(* IEC 61131-3 sources: test/Class/SafetyBaseFSoE (part 5) *)

      pSafetyManagerThis^.NewInst(#MyPara, #MyResult);

      QuitComError := MyResult.aData[0]$DINT;

      // refresh the server on the outer object
      RefreshAsySrv();
    end_if;

    // if we are reinitializing and we have a valid safety number
    if (SafetyState = _ReinitConfig) & SafetyNumber then

      // check every 3 seconds if the cpu is configured
      if b_CheckConfigured & ((ops.tAbsolute - ud_LastCheckConfig) > 3000) then

        // get state via SDO communication
        sd_retval := SDOStdRequ ( us_Command      := SBF_SDO_COMMAND_GET_STATE
                                , p_us_RespData   := ( #GetStateResp )$^USINT
                                , us_RespLength   := sizeof(GetStateResponseType)
                                );

        // the cpu is configured, load the new configuration
        if ( sd_retval = 0 ) &
           (GetStateResp.ConfigState <> SBF_CFG_STATE_UNKNOWN) &
           (GetStateResp.ConfigState <> SBF_CFG_STATE_INVALID) &
           (GetStateResp.ConfigState <> SBF_CFG_STATE_NOT_CONFIGURED) then

          b_CheckConfigured := FALSE;

          b_GetNewConfiguration := TRUE;
        end_if;

        // remember the last time we checked for configurated cpu
        ud_LastCheckConfig := ops.tAbsolute;
      end_if;

      // if there is a new configuration => get it
      if b_GetNewConfiguration then
        // get configuration from safe CPU and build routing tables
        sd_retval := GetRoutingData();
        if sd_retval = 0 then
          b_GetNewConfiguration := FALSE;

          SendAllUnsafeValues();
        else
          LogError("@024B (SafetyBaseFSoE::Background) FAILED TO REINIT THE SAFECPU: .");
        end_if;
      end_if;
    elsif ConnectionInfos.ConnectionNo then
      // if there are still connections => check if they are initialized
      CheckFSoEConnections();
    end_if;

    // here we save the log file from the module to the harddrive (started by user)
    if DiagVars.SavingLogInProgress then

      case DiagVars.SavingLogSSW of

  // ********************************************************************************************************************************************
        GetLogHeader:     // get log header from module (contains size of log memory and write counter)

          // get log header via SDO communication
          sd_retval := SDORequ ( us_Command      := SBF_SDO_COMMAND_GET_LOG_HDR
                               , p_us_RequData   := #DiagVars.ucChoiceSaveLog
                               , us_RequLength   := 1
                               , p_us_RespData   := ( #DiagVars.LogHeader)$^USINT
                               , us_RespLength   := sizeof(DiagStructType.LogHeader)
                               );

          if ( sd_retval = 0 ) then
            DiagVars.LogMemToGet := DiagVars.LogHeader.LogMemSize;
            DiagVars.pLogFileMem$pVoid := ToStdLib.Malloc(size:=DiagVars.LogHeader.LogMemSize);
            //_memset(dest:=DiagVars.pLogFileMem$pVoid, usByte:=0, cntr:=DiagVars.LogHeader.LogMemSize);
            if DiagVars.ucChoiceSaveLog = 0 then
              DiagVars.ReadBaseAdr := SBF_SDO_ADDRESS_LOG_UC1;
            else
              DiagVars.ReadBaseAdr := SBF_SDO_ADDRESS_LOG_UC2;
            end_if;
            DiagVars.SavingLogSSW := GetLogFileBlocks;

          end_if;

  // ********************************************************************************************************************************************
        GetLogFileBlocks: // get the log memory from the application memory of the module (every cycle only a little bit to prevent runtime error in module)

          // we wait here until UpdateCy finishes our work

  // ********************************************************************************************************************************************
        GetLogHeader2:    // get log header from module again. if write counter changed,
                          // we repeat GetLogFileBlocks. otherwise we continue to save the file

          LastWriteCounter := DiagVars.LogHeader.WriteCounter;

          // get LogHeader
          sd_retval := SDORequ ( us_Command      := SBF_SDO_COMMAND_GET_LOG_HDR
                               , p_us_RequData   := #DiagVars.ucChoiceSaveLog
                               , us_RequLength   := 1
                               , p_us_RespData   := ( #DiagVars.LogHeader)$^USINT
                               , us_RespLength   := sizeof(DiagStructType.LogHeader)
                               );

          if ( sd_retval = 0 ) then

            // if write counter is different, repeat last step
            if DiagVars.LogHeader.WriteCounter <> LastWriteCounter then
              DiagVars.SavingLogSSW := GetLogFileBlocks;

              DiagVars.LogMemToGet := DiagVars.LogHeader.LogMemSize;

              // realloc memory (maybe it's a different size)
              ToStdLib.Free(mptr:=DiagVars.pLogFileMem$pVoid);
              DiagVars.pLogFileMem$pVoid := ToStdLib.Malloc(size:=DiagVars.LogHeader.LogMemSize);
            else
              // write counter is equal. continue to last step
              DiagVars.SavingLogSSW := SaveLogFile;
            end_if;
          end_if;

  // ********************************************************************************************************************************************
        SaveLogFile:      // save the memory to the specified file (DPNE)

          // open file (create/overwrite always)
          FileHandle := FileSys.FileOpen(filename:=#DiagVars.DPNE[0], attributes:=ATT_CREATE_ALWAYS);

          DiagVars.SavingLogSuccessful := 1;

          if FileHandle >= 0 then

            // save content to it
            if FileSys.FileWrite(handle:=FileHandle, buffer:=DiagVars.pLogFileMem, length:=DiagVars.LogHeader.LogMemSize) <> DiagVars.LogHeader.LogMemSize$DINT then
              // failed to write to file
              LogError("@024C (SafetyBaseFSoE::Background) Failed to write to binary LogFile.");
              DiagVars.SavingLogSuccessful := -1;
            end_if;

            // close file
            FileSys.FileClose(handle:=FileHandle);
          else
            // failed to open file
            LogError("@024D (SafetyBaseFSoE::Background) Failed to open binary LogFile.");
            DiagVars.SavingLogSuccessful := -1;
          end_if;

          ToStdLib.Free(mptr:=DiagVars.pLogFileMem$pVoid);
          DiagVars.pLogFileMem := NIL;

          DiagVars.SavingLogSSW := GetLogHeader;
          DiagVars.SavingLogInProgress := FALSE;

      end_case;
    end_if;
  end_if;

  state := READY;

END_FUNCTION

FUNCTION VIRTUAL GLOBAL SafetyBaseFSoE::RtWork
  VAR_INPUT
    EAX 	: UDINT;
  END_VAR
  VAR_OUTPUT
    state (EAX) 	: UDINT;
  END_VAR
  VAR
    calloption    : UDINT;
    PDOLength     : UINT;
    pBuffer       : ^USINT;
    pDOInfo       : ^t_DOInfo;
    i             : USINT;
  END_VAR

  // Save state
  // This must be the 1. line in this function or EAX may be overwritten by the generated AWL code
  calloption := EAX;

  if calloption = CALL_OPTION_RT_PRESCAN then    // Called from UpdateRt

//============================ Profiler start======================================================
#ifdef  DM_Profiler
    StartTimeMeasurement(usMode := DMTIME_RT);
#endif
//============================ Profiler end========================================================

    // do pdo communication only, if module has been found and initialized correctly and if there are some LEDs on (else a FW-Update is running)
    if Online &
       (( SafetyState = _SafetyClassOK ) | ( SafetyState = _WaitForSynchronicity ) | ( SafetyState = _ReinitConfig ) | ( SafetyState = _ModFromCfgNotFound ) | ( SafetyState = _UnknownCfgError ) | ( SafetyState = _UnsafeVarNotFound )) then

      // get I/O state, runstate, error
      UpDateNotStd(calloption:=calloption);

      // wait until the safetymanager has initialized everything
      if b_ManagerInitialisationFinished = FALSE then
        return;
      end_if;

      // if any LED is active, then firmware update is not active and we can do our work
      if (VoltageOK | RunState | ServiceMode | ErrorState) then
        // if we are in run state
        if RunState then
          if PDOSingleRunActive & WriteDOsUsed then
            PDOSingleRunActive -= 1;
            if PDOSingleRunActive = 0 then
              for i := 0 to WriteDOsUsed-1 do
                SetDORunState(Handle:=aWritePDOs[i].Handle, NewState:=_BUS_IF_RUN_STATE_NO_RUN);
              end_for;
            end_if;
          end_if;

          //read PDO from hardware, only if PDO is needed by other moduls
          if ( PDOOutputIsUsed ) & ReadDOsUsed then

            PDOLength := pPDOLengthInfoData^.PDOReadLength;

            // only if length is bigger than minimum and smaller than maximum
            if ( PDOLength >= SBF_SPDO_MIN_LENGTH ) & ( PDOLength <= MyPDOReadSize) then

              pBuffer := #PDOOutputBuffer[0];
              pDOInfo := #aReadPDOs[0];
              for i := 0 to (ReadDOsUsed-1) do
                _memcpy(ptr1:=pBuffer, ptr2:=pDOInfo^.pData, cntr:=pDOInfo^.Length);
                pBuffer += pDOInfo^.Length;
                pDOInfo += sizeof(t_DOInfo);
              end_for;

#ifdef SAFETY_PROTOCOL_ANALYZER_ACTIVATED
  RecordFrame(pFrame:=(#PDOOutputBuffer[0])$^DINT, FrameState:=0, IsFSoEPDO:=TRUE);
#endif
            else
              InvalidPDOSizeCnt += 1;
            end_if;
          end_if;
        end_if;
      end_if;
    end_if;

//============================ Profiler start======================================================
#ifdef  DM_Profiler
    StopTimeMeasurement(usMode := DMTIME_RT);
#endif
//============================ Profiler end========================================================

  elsif calloption = CALL_OPTION_RT_POSTSCAN then // Called from UpdateRtPostScan

//============================ Profiler start======================================================
#ifdef  DM_Profiler
    StartTimeMeasurement(usMode := DMTIME_RTPOSTSCAN);
#endif
//============================ Profiler end========================================================

    // do pdo communication only, if module has been found and initialized correctly and if there are some LEDs on (else a FW-Update is running)
    if Online &
       (( SafetyState = _SafetyClassOK ) | ( SafetyState = _WaitForSynchronicity ) | ( SafetyState = _ModFromCfgNotFound ) | ( SafetyState = _UnknownCfgError ) | ( SafetyState = _UnsafeVarNotFound )) then

      // if any LED is active, then firmware update is not active and we can do our work
      if (VoltageOK | RunState | ServiceMode | ErrorState) then

        // write unsafe I/Os
        UpDateNotStd(calloption:=calloption);

        if RunState & ((us_SetBusReadyState = SetBusReadyFinished) | b_ManualQuit) then
          //write PDO to hardware
          if ( ui_cnt_PDOInputBuffer > 0 ) then
            WritePDO2Module();
          end_if;
        end_if;
      end_if;
    end_if;

//============================ Profiler start======================================================
#ifdef  DM_Profiler
    StopTimeMeasurement(usMode := DMTIME_RTPOSTSCAN);
#endif
//============================ Profiler end========================================================
  end_if;

  state := READY;

END_FUNCTION

FUNCTION VIRTUAL GLOBAL SafetyBaseFSoE::ConnectEvent
  VAR
    MyPara 	              : CmdStruct;
    MyResult	            : results;
  END_VAR

  //start DOs
  StartDO();

  if SafetyState = _ModuleNotFound then
    if ModuleSyncNo = 0 then
      SetSafetyState(NewState:=_SafetyClassOK);
    else
      SetSafetyState(NewState:=_WaitForSynchronicity);
    end_if;
  end_if;

  // if we we're already connected => tell the sdias manager we're back (safetythis has to be valid if b_Reconnect is set, therefore we don't have to check it here)
  if b_Reconnect then
    MyPara.uiCmd := CMD_SM_MODULE_RECONNECT;
    MyPara.aPara[0] := THIS$DINT;
    pSafetyManagerThis^.NewInst(#MyPara, #MyResult);
  end_if;

  // whenever the postinit has passed and we got a connect (module has been plugged in after booting the application) => get it's config
  if b_PostInitPassed = TRUE then
    // start reading the config in background (if we're in init the post-init read-out will be faster)

    // next time we check for the configured state of the cpu
    b_CheckConfigured := TRUE;

    // check again in background
    SetSafetyState(NewState:=_ReinitConfig);
  end_if;

// online is set if module init succeeds
//  Online := 1;

END_FUNCTION

FUNCTION VIRTUAL GLOBAL SafetyBaseFSoE::DisconnectEvent
  VAR
    MyPara 	              : CmdStruct;
    MyResult	            : results;
  END_VAR

  //stop DOs
  StopDO();

  // reset time sync state and tell the manager
  if pSafetyManagerThis then
    MyPara.uiCmd := CMD_SM_MODULE_DISCONNECT;
    MyPara.aPara[0] := THIS$DINT;
    pSafetyManagerThis^.NewInst(#MyPara, #MyResult);

    b_Reconnect := TRUE;
  end_if;

  // clear request, otherwise problems could occur on next connect
  LastRequest := _NoOpenRequest;
  ud_AsyComRetryCounter := 0; // reset retry counter

  SafetyNumber := 0;
  FirmwareVersion := 0;

  // increment the config checksum to ensure the readout on reconnect (config readout also contains check of connected modules)
  DesignerPrjConfigCRC += 1;

  SetSafetyState(NewState:=_ModuleNotFound);

  // remove the cpu from all classes, which use it
  ResetConfig();

  if UnsafeScheduler <> UnsafeSchedulerSetBusReady then
    us_SetBusReadyState := WaitPDOsSyncron;
    UnsafeScheduler := UnsafeSchedulerSetBusReady;
  end_if;

  MaxVarsPerReadPackage := 0;
  ReadFramesNeeded := 0;
  MaxVarsPerWritePackage := 0;
  WriteFramesNeeded := 0;

  Online := 0;

END_FUNCTION

FUNCTION VIRTUAL GLOBAL SafetyBaseFSoE::InterruptEvent

END_FUNCTION

FUNCTION SafetyBaseFSoE::SetDORunState
  VAR_INPUT
    Handle 	: UDINT;
    NewState 	: t_BusIFRunState;
  END_VAR
  VAR
    dataSETRUNSTATE : t_SetRunStateCfg;
    tempCmd : CmdStruct;
    _result : results;
  END_VAR

  // set runstate of read
  dataSETRUNSTATE.Handle      := Handle;
  dataSETRUNSTATE.NewRunState := NewState;

  tempCmd.uiCmd         := _BUS_IF_SET_RUN_STATE;
  tempCmd.aPara[0]      := (#dataSETRUNSTATE)$DINT;

  ToBusInterface.NewInst(pPara:=#tempCmd, pResult:=#_result);

  if _result.aData[0]$t_BusIFRetvalErrorcode <> _BUS_IF_RETVAL_OK then
    if NewState = _BUS_IF_RUN_STATE_NO_RUN then
      DOStopFailCounter += 1;
    else
      DOStartFailCounter += 1;
    end_if;
  end_if;

END_FUNCTION

FUNCTION VIRTUAL GLOBAL SafetyBaseFSoE::CyWork
  VAR_INPUT
    EAX 	: UDINT;
  END_VAR
  VAR_OUTPUT
    state (EAX) 	: UDINT;
  END_VAR
  VAR
    p_SDO_act             : ^SDOHeader;
    us_SDO_length         : USINT;
    i                     : UINT;
    p_ReceiveObj          : pVirtualBase;
    p_SDOviaPath          : ^SDOviaPath;
    sd_retval             : DINT;
    IsStandardResp        : BOOL;
    SDORequestBuffer      : SDORequReadConfig;
    DataLen               : USINT;
    us_UnsafeSchedulerRun : USINT;
    p_PDOInBufferAct      : ^PDOInputBuffer;
    EverythingSynchron    : BOOL;
    MyPara 	              : CmdStruct;
    MyResult	            : results;
    UnsafeWrPackageNo     : USINT;
    aUnsafeWrPackages     : UnsafeWritePackages;
    UnsafeRdPackageNo     : USINT;
    aUnsafeRdPackages     : UnsafeReadPackages;
    TmpVal                : DINT;
    AddUnsafePackage      : BOOL;
    GotNewUnsafeValue     : BOOL;
    pHelpUnsafe           : ^UnsafeIORoutingElement;
    BDINTWriteVars        : USINT;
    pAddDynSlaveResp      : ^t_AddDynSlaveResponse;
  END_VAR

//============================ Profiler start======================================================
#ifdef  DM_Profiler
  StartTimeMeasurement(usMode := DMTIME_CY);
#endif
//============================ Profiler end========================================================

#ifdef HWK_SHOW_PRAGMA_MESSAGES
  if b_LogFirstDone = 1 then
    for i := 0 to (ui_cnt_PDOInputBuffer-1) do
      LogValue("@027F (SafetyBaseFSoE::WritePDO2Module) Copy 0x{0} Bytes to offset 0x{1} of Write PDO Nr. 0x{2}", Value:=aLogValues[i].ByteLen, Value2:=aLogValues[i].Offset, Value3:=aLogValues[i].DOIndex);
    end_for;

    b_LogFirstDone := 2;
  end_if;
#endif

  // do sdo communication only, if module has been found and initialized correctly and if there are some LEDs on (else a FW-Update is running)
  if Online & (VoltageOK | RunState | ServiceMode | ErrorState) &
     (( SafetyState <> _ModuleNotFound ) & ( SafetyState <> _MemAllocFailed ) & ( SafetyState <> _LostPowerSupply ) & ( SafetyState <> _ReadFWVerFailed ) & ( SafetyState <> _WrongSafetyHW ) & ( SafetyState <> _ReinitConfig )) then

    // wait until the safetymanager has initialized connection
    if (b_ManagerReadyForSDO = FALSE) then
      return;
    end_if;

    //Update of service messages doesn't take place in realtime

    //read SDO from module and send it to the target module
    //check, if SDO is available and valid
    if ( p_Handle_SDO_Read^.us_Status = SAFETY_SDO_DATA_VALID ) then

      //calculate length of SDO
      us_SDO_length := sizeof(SDOHeader.StdHeader.CRC) + p_Handle_SDO_Read^.SDOStructure.SDOHeader.StdHeader.Len;

      //copy SDO without first byte (=status byte)
      ToStdLib.MemCpy(dest := p_SDOOutputBuffer, source := #p_Handle_SDO_Read^.SDOStructure, size := us_SDO_length );

#ifdef SAFETY_PROTOCOL_ANALYZER_ACTIVATED
  RecordFrame(p_SDOOutputBuffer$^DINT, 0);
#endif

      //mark data as received
      p_Handle_SDO_Read^.us_Status := SAFETY_SDO_NO_DATA;

      //find target object for routing
      p_ReceiveObj := NIL;

      IsStandardResp := FALSE;
      //check, if receiver is addressed by safety number or hardware path
      if ((p_SDOOutputBuffer^.SDOHeader.StdHeader.Typ$USINT AND SBF_SSDO_MASK_TYPE)$t_SafetyFrameType = SSDO_MOD) then

        //search this-pointer of receiver with safety number
        p_ReceiveObj := ( GetRoutingPointerByNumber(ud_SafeNumber := p_SDOOutputBuffer^.SDOHeader.DstAdr))$pVirtualBase;

      elsif ((p_SDOOutputBuffer^.SDOHeader.StdHeader.Typ$USINT AND SBF_SSDO_MASK_TYPE)$t_SafetyFrameType = SSDO_MOD_TP) then

        //search this-pointer of receiver with hardware path
        p_SDOviaPath := p_SDOOutputBuffer$^SDOviaPath;
        p_ReceiveObj := ( GetRoutingPointerByPath(p_ActObjectPath := #p_SDOviaPath^.TopologyPath[0], p_SDOviaPath^.StdHeader.Len - 8))$pVirtualBase;
      elsif ((p_SDOOutputBuffer^.SDOHeader.StdHeader.Typ$USINT AND SBF_SSDO_MASK_TYPE)$t_SafetyFrameType = SDO_STD) then
        IsStandardResp := TRUE;
        StandardResponse := (p_SDOOutputBuffer$^StandardFrameType)^;
        if StandardResponse.SDOHeader.SeqNr = (StandardSeqNr OR 16#80) then

          // if the microcontroller got powered again and we have an SDO response => also get the configuration (don't wait the whole time)
          //if b_WaitForFirmwareBoot = TRUE then // no if to be faster (if it's false, it does not matter if we set it again to false)
          b_WaitForFirmwareBoot := FALSE;
          //end_if;

          case LastRequest of
            _NoOpenRequest: // error, no open request, but we got a response
              LogError("@0252 (SafetyBaseFSoE::CyWork) Standard frame response received, without open request.");

            _SetBusReady:
              IF StandardResponse.SDOHeader.Cmd = SBF_SDO_COMMAND_SET_BUS_READY THEN
                if us_SetBusReadyState <> SendSetBusReady then
                  LogError("@0253 (SafetyBaseFSoE::CyWork) Got Response of SetBusReady, but SSW is not in the right step.");
                  return;
                end_if;
                us_SetBusReadyState := SetBusReadyFinished;
                b_ManualQuit := FALSE;
                UnsafeScheduler := UnsafeSchedulerGetDiagVars; // Go on with the action-steps, done here so we don't lose a whole cycle
                LastRequest := _NoOpenRequest;
                ud_AsyComRetryCounter := 0; // reset retry counter
                if SafetyState = _WaitForSynchronicity then
                  SetSafetyState(NewState:=_SafetyClassOK);
                end_if;
              else
                LogError("@0256 (SafetyBaseFSoE::CyWork) Invalid command: bus ready expected.");
              END_IF;

            _ReadData:
              // if we did read command, then save the value to corresponding server
              if StandardResponse.SDOHeader.Cmd = SBF_SDO_COMMAND_READ then
                // if returncode is 0 read succeeded
                if StandardResponse.aData[0] = 0 then
                  // check if length is correct
                  if StandardResponse.aData[1] = StandardRequest.aData[4] then
                    // delete request
                    LastRequest := _NoOpenRequest;
                    ud_AsyComRetryCounter := 0; // reset retry counter

                    if (DiagVars.SavingLogSSW = GetLogFileBlocks) then
                      // save the last block in the memory for the file
                      _memcpy(ptr1:=DiagVars.pLogFileMem$pVoid + (DiagVars.LogHeader.LogMemSize - DiagVars.LogMemToGet),
                              ptr2:=#StandardResponse.aData[2],
                              cntr:=DiagVars.BytesToGet);

                      DiagVars.LogMemToGet -= DiagVars.BytesToGet;

                      if DiagVars.LogMemToGet = 0 then
                        DiagVars.SavingLogSSW := GetLogHeader2;
                      end_if;
                    else
                      LogError("@0255 (SafetyBaseFSoE::CyWork) SDO Receive: Invalid Read response (no diagnostic read active).");
                    end_if;
                  end_if;
                end_if;
              else
                LogError("@0256 (SafetyBaseFSoE::CyWork) SDO Receive: Invalid command, read expected.");
              end_if;

            _ReadValues:
              // if we did read command, then save the value to corresponding server
              if StandardResponse.SDOHeader.Cmd = SBF_SDO_COMMAND_READ_VALUES then
                // if returncode is 0 read succeeded
                if StandardResponse.aData[0] = 0 then
                  // check if length is correct
                  if StandardResponse.aData[1] = StandardRequest.aData[0] then
                    // delete request
                    LastRequest := _NoOpenRequest;
                    ud_AsyComRetryCounter := 0; // reset retry counter

                    // if we got some outputs in the routing table and a valid pointer, write values to servers
                    if ui_CntUnsafeOutputs & pUnsafeOutElement then

                      // depending on length we do different number of server write-methods to set the data we just read
//                      pUnsafeOutElement := p_UnsafeOutputsTable + (UnsafeReadTransNr * MaxVarsPerReadPackage * sizeof(UnsafeIORoutingElement));  // the pointer is already on this element
                      for i := 0 to (StandardResponse.aData[1] - 1) do
                        // save the new value temporarily
                        TmpVal := StandardResponse.aData[2 + (i * sizeof(DINT))]$DINT;
                        if pUnsafeOutElement^.ud_Thisp then
                          if pUnsafeOutElement^.UnsafeType = BDINTOutput then
                            pUnsafeOutElement^.sd_OldValue := RD(pUnsafeOutElement^.ud_Thisp$^void)$DINT;
                            TmpVal := ((pUnsafeOutElement^.sd_OldValue$UDINT AND (NOT pUnsafeOutElement^.BitMask)) OR
                                      (TmpVal$UDINT AND pUnsafeOutElement^.BitMask))$DINT;

                            // now we have to write the value to the server
                            WR(pUnsafeOutElement^.ud_Thisp$^void, TmpVal);
                          else
                            WR(pUnsafeOutElement^.ud_Thisp$^void, TmpVal);
                          end_if;
                        elsif (pUnsafeOutElement^.UnsafeType = ExternalOutput) | (pUnsafeOutElement^.UnsafeType = ExternalBDINTOutput) then
                          pUnsafeOutElement^.sd_NewValue4External := TmpVal;

                          // mark the value as valid
                          pUnsafeOutElement^.b_IsValid := TRUE;
                        end_if;
                        pUnsafeOutElement += sizeof(UnsafeIORoutingElement);
                      end_for;
                    end_if;

                    UnsafeReadTransNr += 1;
                  end_if;
                end_if;
              else
                LogError("@0257 (SafetyBaseFSoE::CyWork) SDO Receive: Invalid command, read values expected.");
              end_if;

            _WriteValues:
              if IsOptimizedCPU() then
                // if we did a write command, just check
                if StandardResponse.SDOHeader.Cmd = SBF_SDO_COMMAND_WRITE_VALUES then
                  // delete request
                  LastRequest := _NoOpenRequest;
                  ud_AsyComRetryCounter := 0; // reset retry counter

                  // if there is no more element to send or check for changes => proceed to the next step
                  if pUnsafeInElement = NIL then
                    UnsafeScheduler := UnsafeSchedulerReadData; //We need to set scheduler to next step....
                  end_if;
                else
                  LogError("@0258 (SafetyBaseFSoE::CyWork) SDO Receive: Invalid command, write expected.");
                end_if;
              else
                // on CSCP011 the SDO_COMMAND_WRITE_VALUES didn't exist

                // if we did a write command, just check
                if StandardResponse.SDOHeader.Cmd = SBF_SDO_COMMAND_WRITE then
                  // delete request
                  LastRequest := _NoOpenRequest;
                  ud_AsyComRetryCounter := 0; // reset retry counter

                  if UnsafeWriteTransNr < (WriteFramesNeeded - 1) then
                    UnsafeWriteTransNr += 1;
                  else
                    UnsafeWriteTransNr := 0;
                    UnsafeWritingActive := FALSE;
                    UnsafeScheduler := UnsafeSchedulerReadData; //We need to set scheduler to next step....
                  end_if;
                else
                  LogError("@0258 (SafetyBaseFSoE::CyWork) SDO Receive: Invalid command, write expected.");
                end_if;
              end_if;

            _GetCRC:
              // check if it's a response to a read command
              if StandardResponse.SDOHeader.Cmd = SBF_SDO_COMMAND_READ then
                // if returncode is 0 read succeeded
                if StandardResponse.aData[0] = 0 then
                  // check if length is correct
                  if StandardResponse.aData[1] = 4 then

                    // delete request
                    LastRequest := _NoOpenRequest;
                    ud_AsyComRetryCounter := 0; // reset retry counter

                    if DesignerPrjConfigCRC <> StandardResponse.aData[2]$UDINT then
                      // CRC has changed => save the new crc
                      DesignerPrjConfigCRC := StandardResponse.aData[2]$UDINT;

                      // show that we read the config of the class again
                      SetSafetyState(NewState:=_ReinitConfig);

                      if pSafetyManagerThis then
                        MyPara.uiCmd := CMD_SM_NEW_SAFETY_PROJECT;
                        MyPara.aPara[0] := 4;
                        MyPara.aPara[4] := (#SafetyNumber)$DINT;
                        pSafetyManagerThis^.NewInst(#MyPara, #MyResult);
                      end_if;

                      // remove the cpu from all classes, which use it
                      ResetConfig();

                      // we have to return here because:
                      // the command CMD_SM_NEW_SAFETY_PROJECT will trigger a disconnect of this class which will set the unsafe scheduler to setbusready,
                      // which would skip the synchron check in the actual cyclic run because everything of the old configuration is synchron now
                      return;
                    end_if;
                  end_if;
                end_if;
              end_if;

            _WriteSysTime:
              if StandardResponse.SDOHeader.Cmd = SBF_SDO_COMMAND_WRITE then
                // if returncode is 0 read succeeded
                if StandardResponse.aData[0] = 0 then
                  // delete request
                  LastRequest := _NoOpenRequest;
                  ud_AsyComRetryCounter := 0; // reset retry counter
                end_if;
              else
                LogError("@0258 (SafetyBaseFSoE::CyWork) SDO Receive: Invalid command, write expected.");
              end_if;

            _WriteFlexConCommand:
              if StandardResponse.SDOHeader.Cmd = SBF_SDO_COMMAND_WRITE then
                // if returncode is 0 read succeeded
                if StandardResponse.aData[0] = 0 then
                  // delete request
                  LastRequest := _NoOpenRequest;
                  ud_AsyComRetryCounter := 0; // reset retry counter
                end_if;
              else
                LogError("@0258 (SafetyBaseFSoE::CyWork) SDO Receive: Invalid command, write expected.");
              end_if;

            _DiagState:
              if StandardResponse.SDOHeader.Cmd = SBF_SDO_COMMAND_GET_STATE then
                _memcpy(ptr1 := #DiagVars.UserGetStateResp,
                        ptr2 := #StandardResponse.aData + SIZEOF(USINT),
                        cntr := sizeof(GetStateResponseType) );
                DiagVars.UserDiagStateReady := TRUE;
                DiagVars.UserWantsDiagState := FALSE;
                LastRequest := _NoOpenRequest;
                ud_AsyComRetryCounter := 0; // reset retry counter
              end_if;
            _DiagInfo:
              if StandardResponse.SDOHeader.Cmd = SBF_SDO_COMMAND_GET_DIAG_INFO then
                _memcpy(ptr1 := #DiagVars.UserGetDiagInfoResp,
                        ptr2 := #StandardResponse.aData + SIZEOF(USINT),
                        cntr := sizeof(SafetyDiagInfo) );
                DiagVars.UserDiagInfoReady := TRUE;
                DiagVars.UserWantsDiagInfo := FALSE;
                LastRequest := _NoOpenRequest;
                ud_AsyComRetryCounter := 0; // reset retry counter
              end_if;

            _ReadRetryCounter:
              //if we did read command, then save the value to corresponding server
              if StandardResponse.SDOHeader.Cmd = SBF_SDO_COMMAND_READ then
                // if returncode is 0 read succeeded
                if StandardResponse.aData[0] = 0 then
                  // check if length is correct
                  if StandardResponse.aData[1] = SBF_SDO_LENGTH_RETRY_COUNTER then
                    // delete request
                    LastRequest := _NoOpenRequest;
                    ud_AsyComRetryCounter := 0; // reset retry counter

                    //Only Write if Retry Counter has changed
                    if StandardResponse.aData[2] <> us_OldRetryCounter then
                      //if retry counter has changed, save the new retry counter
                      SafetyRetryCounter += to_usint(StandardResponse.aData[2] - us_OldRetryCounter);
                      us_OldRetryCounter := StandardResponse.aData[2];

                      //0x20400000 is adress of retry counter: 1 byte amount of all retries of all modules, 16byte µC1, 16 byte µC2
                      //Save the values from the modules
                      ToStdLib.MemCpy(dest:=#a_RetryCnt[0], source:=#StandardResponse.aData[3], size:=SBF_SDO_LENGTH_RETRY_COUNTER);

                      //Calls the method of class sdiassafetymanager
                      SetRetryCounter();
                    end_if;
                  end_if;
                end_if;
              else
                LogError("@0257 (SafetyBaseFSoE::CyWork) SDO Receive: Invalid command, read values expected.");
              end_if;

            _ErrorChannelInfo:
              //if we did read command, then save the value to corresponding server
              if StandardResponse.SDOHeader.Cmd = SBF_SDO_COMMAND_READ then
                // if returncode is 0 read succeeded
                if StandardResponse.aData[0] = 0 then
                  // check if length is correct
                  if StandardResponse.aData[1] <> 0  then
                    _memcpy(ptr1 := #aErrorMem[actoffset],
                            ptr2 := #StandardResponse.aData[2],
                            cntr := StandardResponse.aData[1]);
                    if remainingPacketlength = 0 then
                      remainingPacketlength := StandardResponse.aData[2] - StandardResponse.aData[1];
                      actoffset := StandardResponse.aData[1];
                    else
                      remainingPacketlength -= StandardResponse.aData[1];
                      actoffset += StandardResponse.aData[1];
                    end_if;

                    // delete request
                    LastRequest := _NoOpenRequest;
                    ud_AsyComRetryCounter := 0; // reset retry counter
                    if remainingPacketlength <= 0  then
                      //Finish
                      DiagVars.UserErrorInfoReady := TRUE;
                      DiagVars.UserWantsErrorInfo := FALSE;
                      remainingPacketlength := 0; //reset remainingPacketlength
                      actoffset := 0; //reset offset
                    end_if;
                  end_if;
                end_if;
              end_if;

            _ReadFlexConNodeState:
              //if we did read command, then save the value to corresponding server
              if StandardResponse.SDOHeader.Cmd = SBF_SDO_COMMAND_READ then
                // if returncode is 0 read succeeded
                if StandardResponse.aData[0] = 0 then
                  // check if length is correct
                  if StandardResponse.aData[1] = sizeof(t_FlexConNodeState) then

                    // store the structure locally
                    _memcpy(ptr1 := #sFlexCon.LastNodeState,
                            ptr2 := #StandardResponse.aData[2],
                            cntr := StandardResponse.aData[1]);

                    // save the values to the server of the object
                    sFlexCon.pCommand^            := sFlexCon.LastNodeState.Command;
                    sFlexCon.pStateMachine^       := sFlexCon.LastNodeState.StateMachine;
                    sFlexCon.pHostSafetyNumber^   := sFlexCon.LastNodeState.HostSafetyNumber;

                    // delete request
                    LastRequest := _NoOpenRequest;
                    ud_AsyComRetryCounter := 0; // reset retry counter
                  end_if;
                end_if;
              end_if;

            _ReadFlexConHostState:
              //if we did read command, then save the value to corresponding server
              if StandardResponse.SDOHeader.Cmd = SBF_SDO_COMMAND_READ then
                // if returncode is 0 read succeeded
                if StandardResponse.aData[0] = 0 then
                  // check if length is correct (maximum the requested size)
                  if StandardResponse.aData[1] & (StandardResponse.aData[1] <= sFlexCon.LastHostState.LastRequestedLength) then
                    // if the size in the response is smaller than the requested (we already got everything in the first package)
                    if StandardResponse.aData[1] <= sFlexCon.LastHostState.LastRequestedLength then
                      // adjust the last requested length to the received for correct handling of the received data
                      sFlexCon.LastHostState.LastRequestedLength := StandardResponse.aData[1];
                    end_if;

                    // if it's the first package
                    if sFlexCon.LastHostState.CurrentReadOffset = 0 then
                      // if length is ok and there is at least 1 connection but not more than the maximum
                      if (StandardResponse.aData[1] >= sizeof(HDINT)) & StandardResponse.aData[2]$HDINT & (StandardResponse.aData[2]$HDINT <= MAX_FSOE_CONNECTIONS) then
                        // the first 4 byte contain the number of connections following
                        sFlexCon.LastHostState.NoConnections := StandardResponse.aData[2]$HDINT;
                        _memcpy(ptr1:=#sFlexCon.LastHostState.aConnections[0], ptr2:=#StandardResponse.aData[2] + sizeof(HDINT), cntr:=sFlexCon.LastHostState.LastRequestedLength - sizeof(HDINT));

                        // calculate how many bytes are missing (what do we need minus what do we already have)
                        sFlexCon.LastHostState.BytesMissing       := sFlexCon.LastHostState.NoConnections$UINT * sizeof(HDINT) + sizeof(HDINT) - sFlexCon.LastHostState.LastRequestedLength;
                        sFlexCon.LastHostState.CurrentReadOffset  += sFlexCon.LastHostState.LastRequestedLength;
                      else
                        // no connection or too many to fit into the array
                        sFlexCon.LastHostState.NoConnections := 0;

                        // nothing missing
                        sFlexCon.LastHostState.BytesMissing := 0;
                      end_if;
                    else
                      // offset is not zero => follow up package
                      _memcpy(ptr1:=#sFlexCon.LastHostState.aConnections[0] + sFlexCon.LastHostState.CurrentReadOffset - sizeof(HDINT), ptr2:=#StandardResponse.aData[2], cntr:=sFlexCon.LastHostState.LastRequestedLength);

                      // update the bytes missing and the current reading offset
                      sFlexCon.LastHostState.BytesMissing      -= sFlexCon.LastHostState.LastRequestedLength;
                      sFlexCon.LastHostState.CurrentReadOffset += sFlexCon.LastHostState.LastRequestedLength;
                    end_if;
                  else
                    // wrong length => reset number of connections
                    sFlexCon.LastHostState.NoConnections := 0;

                    // nothing missing
                    sFlexCon.LastHostState.BytesMissing := 0;
                  end_if;

                  // if we got all data
                  if sFlexCon.LastHostState.BytesMissing = 0 then

                    // update connection state at managing modules
                    MyPara.uiCmd := CMD_SM_UPDATE_FLEX_CON_HOST;
                    MyPara.aPara[0] := sFlexCon.LastHostState.NoConnections$DINT;
                    MyPara.aPara[1] := (#sFlexCon.LastHostState.aConnections[0])$DINT;
                    pSafetyManagerThis^.NewInst(#MyPara, #MyResult);

                    // reset the offset so we start reading at 0 in the next round
                    sFlexCon.LastHostState.CurrentReadOffset := 0;

                    // reset timemark
                    sFlexCon.ud_LastHostStateTimeStamp := ops.tAbsolute;
                  end_if;

                  // delete request
                  LastRequest := _NoOpenRequest;
                  ud_AsyComRetryCounter := 0; // reset retry counter

                end_if;
              end_if;

          else
            LogError("@025A (SafetyBaseFSoE::CyWork) SDO Receive: Invalid standard frame response.");
          end_case;

          // if request is deleted, increase sequence number to set next request
          if LastRequest = _NoOpenRequest then
            if StandardSeqNr < 16#7F then
              StandardSeqNr += 1;
            else
              StandardSeqNr := 0;
            end_if;
          end_if;
        else
          LogError("@025B (SafetyBaseFSoE::CyWork) SDO Receive: Invalid sequence number in Standard SDO response.");
          LogValue("expected: 0x{0} / received: 0x{1}", Value:=(StandardSeqNr OR 16#80), Value2:=StandardResponse.SDOHeader.SeqNr);
        end_if;
      elsif ((p_SDOOutputBuffer^.SDOHeader.StdHeader.Typ$USINT AND SBF_SSDO_MASK_TYPE)$t_SafetyFrameType = SSDO_MOD_DEVADDR) then

        //Check if we know our target
        p_ReceiveObj := ( GetRoutingPointerByNumber(ud_SafeNumber := p_SDOOutputBuffer^.SDOHeader.DstAdr))$pVirtualBase;

        //Forward data to manager if we found no routing target, otherwise the SDO will be directly send to target
        if p_ReceiveObj = NIL then

          // Forward to manager if possible
          if pSafetyManagerThis & us_SDO_length then
  #ifdef DO_DEBUG
            DOCheck(pFrame:=(p_SDOOutputBuffer)$^t_SDOStdHeader, pCheckStruct:=#SDORead);
  #endif

            if ( (p_SDOOutputBuffer^.SDOHeader.StdHeader.Cmd = SBF_SDO_COMMAND_ADD_DYN_SLAVE) | (p_SDOOutputBuffer^.SDOHeader.StdHeader.Cmd = SBF_SDO_COMMAND_ADD_DYN_SLAVE2) )&
               (p_SDOOutputBuffer^.SDOHeader.StdHeader.Typ$USINT AND SBF_SSDO_MASK_RESPONSE) then
              // we need a response big enough to hold our info, the returncode must be 0 and the offset/length info has to be plausible
              if ((p_SDOOutputBuffer^.SDOHeader.StdHeader.Len + sizeof(SDOHeader.StdHeader.CRC)) >= sizeof(t_AddDynSlaveResponse)) &
                  (p_SDOOutputBuffer^.us_Returncode = 0) & CheckAddDynSlaveResponse(p_SDOOutputBuffer$^t_AddDynSlaveResponse) then

                pAddDynSlaveResp := p_SDOOutputBuffer$^t_AddDynSlaveResponse;

                MyPara.aPara[2]       := THIS$DINT;

                MyPara.aPara[3]$HDINT := pAddDynSlaveResp^.OffsetSafeOutData; // offset to data from module
                MyPara.aPara[4]$HDINT := pAddDynSlaveResp^.LenSafeOutData;    // size of data from module

                MyPara.aPara[5]$HDINT := pAddDynSlaveResp^.OffsetSafeInData;  // offset to data to module
                MyPara.aPara[6]$HDINT := pAddDynSlaveResp^.LenSafeInData;     // size of data to module
              else
                _memset(dest:=#MyPara.aPara[2], usByte:=0, cntr:=5*sizeof(DINT));
              end_if;
            end_if;

            MyPara.uiCmd := CMD_SM_SDO_TO_MANAGER;
            MyPara.aPara[0] := to_dint(us_SDO_length);
            MyPara.aPara[1] := p_SDOOutputBuffer$DINT;
            pSafetyManagerThis^.NewInst(#MyPara, #MyResult);

            IsStandardResp := TRUE;
          else
            //log not routable SDOs
            LogValue("@025E (SafetyBaseFSoE::CyWork) Safety module 0x{0}: SDO not routed to receiver {1}", SafetyNumber$UDINT, p_SDOOutputBuffer^.SDOHeader.DstAdr$UDINT);
          end_if;
        end_if;
      else
        LogError("@025C (SafetyBaseFSoE::CyWork) SDO Receive: Invalid frametype in Standard SDO response.");
      end_if;

      //if there is no object, the message will be lost
      if ( p_ReceiveObj ) then

        //send SDO to receiver object
        MyPara.uiCmd := CMD_SM_ADD_SDO_TO_BUFFER;
        MyPara.aPara[0] := p_SDOOutputBuffer$DINT;
        MyPara.aPara[1] := us_SDO_length;
        sd_retval$iprStates := p_ReceiveObj^.NewInst(#MyPara, #MyResult);

//        sd_retval := p_ReceiveObj^.AddSDOToBuffer(p_us_Message := p_SDOOutputBuffer$^USINT, us_length := us_SDO_length);

        if sd_retval$iprStates = ERROR then
          // generate error message with returncode (add to logfile and debugger trace)
          LogValue("@025D (SafetyBaseFSoE::CyWork) AddSDOToBuffer failed: Returncode: -0x{0}", Value:=(0-sd_retval)$UDINT);
        end_if;

      elsif IsStandardResp = FALSE then

        if pSafetyManagerThis & us_SDO_length then
#ifdef DO_DEBUG
          DOCheck(pFrame:=(p_SDOOutputBuffer)$^t_SDOStdHeader, pCheckStruct:=#SDORead);
#endif

          // if the command is get safety number and the compressed path type is 2, it can only be in this system (no interface frame) and therefore forwarding to the manager would not make sense (the class should already find the other module with GetRoutingPointerByPath()
          if (p_SDOOutputBuffer^.SDOHeader.StdHeader.Cmd = SBF_SDO_COMMAND_GET_SAFENBR) &
             (p_SDOOutputBuffer^.SDOHeader.StdHeader.Typ = SSDO_MOD_TP) &
             (p_SDOOutputBuffer^.SDOHeader.DstAdr$USINT = 2) then
            // skip forwarding in this case
          else
            // forward it to the safety manager
            MyPara.uiCmd := CMD_SM_SDO_TO_MANAGER;
            MyPara.aPara[0] := to_dint(us_SDO_length);
            MyPara.aPara[1] := p_SDOOutputBuffer$DINT;
            pSafetyManagerThis^.NewInst(#MyPara, #MyResult);
          end_if;
        else
          //log not routable SDOs
          LogValue("@025E (SafetyBaseFSoE::CyWork) Safety module 0x{0}: SDO not routed to receiver {1}", SafetyNumber$UDINT, p_SDOOutputBuffer^.SDOHeader.DstAdr$UDINT);
        end_if;
      end_if;

    elsif (LastRequest <> _NoOpenRequest) & (ud_TransfertimePerPackage > 0) then
      // count up for timeout
      ud_UnsafeTimeoutCounter += 1;

      if ( ud_UnsafeTimeoutCounter ) > ( 50 * ud_TransfertimePerPackage ) then
        CASE UnsafeScheduler OF

          UnsafeSchedulerSetBusReady:
            LogError("@025F (SafetyBaseFSoE::UpdateCy) Timeout on setting bus ready.");

          UnsafeSchedulerGetDiagVars:
            IF LastRequest = _ReadData THEN
              LogError("@0260 (SafetyBaseFSoE::UpdateCy) Timeout requesting DiagVars.");
            END_IF;
            UnsafeScheduler := UnsafeSchedulerNonPriorData;
            DiagVars.SavingLogSSW := GetLogFileBlocks;

          UnsafeSchedulerNonPriorData:
            if LastRequest = _WriteSysTime then
              LogError("@0497 (SafetyBaseFSoE::UpdateCy) Timeout writing the system time to module.");
            else
              LogError("@0261 (SafetyBaseFSoE::UpdateCy) Timeout requesting CRC.");
            end_if;

            UnsafeScheduler := UnsafeSchedulerWriteData;

          UnsafeSchedulerWriteData:
            LogError("@0262 (SafetyBaseFSoE::UpdateCy) Timeout writing Data 'Unsafe Input'.");
            UnsafeScheduler := UnsafeSchedulerReadData;
            UnsafeWriteTransNr := 0;

          UnsafeSchedulerReadData:
            LogError("@0263 (SafetyBaseFSoE::UpdateCy) Timeout reading Data 'Unsafe Output'.");
            UnsafeScheduler := UnsafeSchedulerDiagState;
            UnsafeReadTransNr := 0;

          UnsafeSchedulerDiagState:
            LogError("@0264 (SafetyBaseFSoE::UpdateCy) Timeout on reading DiagState.");
            UnsafeScheduler := UnsafeSchedulerDiagInfo;

          UnsafeSchedulerDiagInfo:
            LogError("@0265 (SafetyBaseFSoE::UpdateCy) Timeout on reading DiagInfo.");
            UnsafeScheduler := UnsafeSchedulerGetRetryCounter;

          UnsafeSchedulerGetRetryCounter:
            LogError("@0266 (SafetyBaseFSoE::UpdateCy) Timeout on reading RetryCounter.");
            UnsafeScheduler := UnsafeSchedulerChannelError;

          UnsafeSchedulerChannelError:
            LogError("@0267 (SafetyBaseFSoE::UpdateCy) Timeout on reading ChannelErrorInfo.");
            UnsafeScheduler := UnsafeSchedulerGetFlexConNodeState;

          UnsafeSchedulerGetFlexConNodeState:
            LogError("@0267 (SafetyBaseFSoE::UpdateCy) Timeout on reading FlexConNodeState.");
            UnsafeScheduler := UnsafeSchedulerGetFlexConHostState;

          UnsafeSchedulerGetFlexConHostState:
            LogError("@0267 (SafetyBaseFSoE::UpdateCy) Timeout on reading FlexConHostState.");
            UnsafeScheduler := UnsafeSchedulerGetDiagVars;

        END_CASE;

        // we only increase the retry counter if the module is running
        if RunState then
          ud_AsyComRetryCounter += 1;
        end_if;

        if ud_AsyComRetryCounter >= SBF_SDO_MAX_TRIES then
          SetSafetyState(NewState:=_AsyncComError);
          LogError("@0268 (SafetyBaseFSoE::UpdateCy) Too many consecutive asynchronous commands failed! Please contact Sigmatek Support!");
        else
          LastRequest := _NoOpenRequest;
          // if request is deleted, increase sequence number to set next request
          if StandardSeqNr < 16#7F then
            StandardSeqNr += 1;
          else
            StandardSeqNr := 0;
          end_if;
        end_if;
      end_if;

    end_if;

    //write to hardware from other module received SDO
    if ( ui_cnt_SDOInputBuffer > 0 ) & p_SDOInputBuffer then

      //set pointer to first SDO in the SDO list
      p_SDO_act   := p_SDOInputBuffer$^SDOHeader;

      //calculate length of SDO (CRC + data length)
      us_SDO_length := sizeof (SDOHeader.StdHeader.CRC) + p_SDO_act^.StdHeader.Len;

      //check, if buffer is empty
      if ( p_Handle_SDO_Write^.us_Status = SAFETY_SDO_NO_DATA ) then

#ifdef SAFETY_PROTOCOL_ANALYZER_ACTIVATED
  RecordFrame(p_SDO_act$^DINT, 1);
#endif

        //copy SDO into write-buffer
        ToStdLib.MemCpy(dest := #p_Handle_SDO_Write^.SDOStructure, source := p_SDO_act, size := us_SDO_length);

        //mark SDO data as valid
        p_Handle_SDO_Write^.us_Status := SAFETY_SDO_DATA_VALID;

        //decrement amount of SDOs
        ui_cnt_SDOInputBuffer -= 1;

        //if there is at least 1 SDO left, copy the remaining memory over the actual SDO
        if ( ui_cnt_SDOInputBuffer > 0 ) then

          //remove first entry in the SDO list
          _memmove(p_SDOInputBuffer, (p_SDOInputBuffer + SBF_SDO_MAX_LENGTH), (ui_cnt_SDOInputBuffer * SBF_SDO_MAX_LENGTH));
        end_if;
      end_if;
    end_if;

    // if we have to quit the communication errors and there is no other request open at this time
    if (QuitComError = 1) & (LastRequest = _NoOpenRequest) then
      if UnsafeScheduler <> UnsafeSchedulerSetBusReady then
        us_SetBusReadyState := WaitPDOsSyncron;
        UnsafeScheduler := UnsafeSchedulerSetBusReady;
      end_if;

      QuitComError := 0;

      // refresh the server on the outer object
      RefreshAsySrv();
    end_if;

    if ( SafetyState <> _ReinitConfig ) & ( p_Handle_SDO_Write^.us_Status = SAFETY_SDO_NO_DATA ) then

      // priority request before checking the scheduler
      // if the channel is free and we have a command request for the flexible constellation node => send the command
      if (LastRequest = _NoOpenRequest) & (sFlexCon.FoundNodeInConfig) & (sFlexCon.CommandRequest) & b_ManagerInitialisationFinished then

        StandardRequest.SDOHeader.CRC  := 0;                               // CRC is always 0 in Std communication
        StandardRequest.SDOHeader.Cmd  := SBF_SDO_COMMAND_WRITE;           // read command
        StandardRequest.SDOHeader.Typ  := SDO_STD;                         // standard frame type
        StandardRequest.SDOHeader.SeqNr:= StandardSeqNr OR 16#80;          // sequence number
        StandardRequest.SDOHeader.Len  := 4 + 4 + 1 + sizeof(UDINT);       // header + destination address + length of data + size of data
        StandardRequest.aData[0]$UDINT := SBF_SDO_ADDRESS_FLEX_CON_NODE;   // address of the flex con data
        StandardRequest.aData[4]       := sizeof(UDINT);                   // length of data
        StandardRequest.aData[5]$UDINT := sFlexCon.CommandRequest;     // new command

        // reset marker to detect new commands
        sFlexCon.CommandRequest := 0;

        LastRequest := _WriteFlexConCommand;

        //copy SDO into write-buffer
        ToStdLib.MemCpy(dest := #p_Handle_SDO_Write^.SDOStructure, source := #StandardRequest, size := (sizeof(SDOHeader.StdHeader.CRC) + StandardRequest.SDOHeader.Len));

        //mark SDO data as valid
        p_Handle_SDO_Write^.us_Status := SAFETY_SDO_DATA_VALID;

        if ( pISafety^.udVersion >= 16#1001 ) then
          SAFETY_iPushSafetyTask();
        end_if;

      end_if;

      // Start of scheduler; we need to share the time between reading, writing and diagnosis
      us_UnsafeSchedulerRun := 0;

      // number of steps in total minus 1, because the SetBusReady doesn't count here since it's not part of the rotation
      SchedulerStepNo := 10;

      // Check actions until we find somthing we need to do
      // all x (SchedulerStepNo) action-steps must be walked through during one cycle to make sure new data is fetched as fast as possible
      // SetBusReady is an exception: this step is only performed once on bootup!
      while (us_UnsafeSchedulerRun < SchedulerStepNo) & (LastRequest = _NoOpenRequest) do
        us_UnsafeSchedulerRun += 1;
        ud_UnsafeTimeoutCounter := 0; //No active request: we can reset the timeout-counter
        case UnsafeScheduler of
//**********************************************************************************************************************************************************
          UnsafeSchedulerSetBusReady:  // this step is excluded from the rotation (set at startup, on disconnect or quit error)

            //Set Bus Ready has to be done one time after the manager initialisation was finished
            //Other steps of the scheduler can be executed before the manager initialisation is finished (diag steps)
            if b_ManagerInitialisationFinished = TRUE then

              case us_SetBusReadyState of

              //-------------------------------------------------------------------------------------------------------------
                WaitPDOsSyncron:

                  EverythingSynchron := TRUE;

                  // it's possible that all PDOs are coming from a different domain, then we have no inputbuffer
                  if ui_cnt_PDOInputBuffer then
                    p_PDOInBufferAct := #aPDOInputBuffer[0];
                    for i := 0 to (ui_cnt_PDOInputBuffer-1) do
                      if p_PDOInBufferAct^.b_TimeSynchron = FALSE then
                        // we're still not synchron with this module. if it's optional it is probably not connected
                        if p_PDOInBufferAct^.b_IsOptional then
                          if (ops.tAbsolute - ud_OptionalTimeoutStart) <= SBF_OPTIONAL_MODULE_SYNC_TIMEOUT then
                            // if timeout not exceeded => not sychron (otherwise the variable will stay on it's old value)
                            EverythingSynchron := FALSE;
                            exit;
                          else
                            TRACE("Synchronisation timeout for optional module exceeded => assume it's synchon.");
                          end_if;
                        else
                          EverythingSynchron := FALSE;
                          exit;
                        end_if;
                      end_if;

                      p_PDOInBufferAct +=  sizeof(PDOInputBuffer);
                    end_for;

                    if EverythingSynchron & (ModuleSyncNo > 0) then
                      ModuleSyncNo -= 1;

  #ifdef SAFETY_DEBUG_LOGGING_ACTIVATED
  //                  case ud_MyModuleID of
  //                    CSCP01x_ID:
  //                      TRACE("ModuleSyncNo wurde dekrementiert von: CSCP.");
  //
  //                    CSDI16x_ID:
  //                      TRACE("ModuleSyncNo wurde dekrementiert von: CSDI.");
  //
  //                    CSTO08x_ID:
  //                      TRACE("ModuleSyncNo wurde dekrementiert von: CSTO.");
  //                  end_case;
  #endif
                  end_if;
  #ifdef SAFETY_DEBUG_LOGGING_ACTIVATED
  //              elsif EverythingSynchron then
  //                  case ud_MyModuleID of
  //                    CSCP01x_ID:
  //                      TRACE("ModuleSyncNo wurde nicht verändert von: CSCP.");
  //
  //                    CSDI16x_ID:
  //                      TRACE("ModuleSyncNo wurde nicht verändert von: CSDI.");
  //
  //                    CSTO08x_ID:
  //                      TRACE("ModuleSyncNo wurde nicht verändert von: CSTO.");
  //                  end_case;
  #endif
                  end_if;

                  if EverythingSynchron then
                    us_SetBusReadyState := WaitAllModulesSyncron;
                  end_if;

              //-------------------------------------------------------------------------------------------------------------
                WaitAllModulesSyncron:
                  // wait for other modules to be synchron with each other
                  if (ModuleSyncNo = 0) & b_ManagerInitialisationFinished then
                    us_SetBusReadyState := SendSetBusReady;
                  end_if;

              //-------------------------------------------------------------------------------------------------------------
                SendSetBusReady:
                  // send the bus-ready command
                  SDORequestBuffer.StdHeader.CRC  := 0;                                                   // CRC is always 0 in Std communication
                  SDORequestBuffer.StdHeader.Cmd  := SBF_SDO_COMMAND_SET_BUS_READY;                        // set bus ready command
                  SDORequestBuffer.StdHeader.Typ  := SDO_STD;                                             // standard frame type
                  SDORequestBuffer.StdHeader.SeqNr:= StandardSeqNr OR 16#80;                              // sequence number
                  SDORequestBuffer.StdHeader.Len  := 4;                                                   // header

                  LastRequest := _SetBusReady;

  #ifdef SAFETY_PROTOCOL_ANALYZER_ACTIVATED
    RecordFrame((#SDORequestBuffer)$^DINT, 1);
  #endif

                  //copy SDO into write-buffer
                  ToStdLib.MemCpy(dest := #p_Handle_SDO_Write^.SDOStructure, source := #SDORequestBuffer, size := (sizeof(SDOHeader.StdHeader.CRC) + SDORequestBuffer.StdHeader.Len));

                  //mark SDO data as valid
                  p_Handle_SDO_Write^.us_Status := SAFETY_SDO_DATA_VALID;

                  if ( pISafety^.udVersion >= 16#1001 ) then
                    SAFETY_iPushSafetyTask();
                  end_if;

              //-------------------------------------------------------------------------------------------------------------
                SetBusReadyFinished:
                  // all ok, nothing to do here

              end_case;
              us_UnsafeSchedulerRun := 16#FF; //make sure we don't repeat the while-loop until we have sent the bus-ready command

            else
              UnsafeScheduler := UnsafeSchedulerGetDiagVars;  //go on with next step
            end_if;
//**********************************************************************************************************************************************************
          UnsafeSchedulerGetDiagVars:

            //check, if buffer is empty and we got some unsafe data to get/set and crc check is finished
            if (DiagVars.SavingLogSSW = GetLogFileBlocks) then

              // check if more than blocksize to get
              if DiagVars.LogMemToGet > SBF_LOG_DATA_BLOCK_SIZE then
                // get a complete block
                DiagVars.BytesToGet := SBF_LOG_DATA_BLOCK_SIZE;
              else
                // get only the last bytes
                DiagVars.BytesToGet := DiagVars.LogMemToGet$USINT;
              end_if;

              StandardRequest.SDOHeader.Cmd   := SBF_SDO_COMMAND_READ;                         // read command
              StandardRequest.SDOHeader.Typ   := SDO_STD;                                     // standard frame type
              StandardRequest.SDOHeader.SeqNr := StandardSeqNr OR 16#80;                      // sequence number is in special area
              StandardRequest.SDOHeader.Len   := 4 + 4 + 1;                                   // header + destination address + length of data
              StandardRequest.aData[0]$UDINT  := DiagVars.ReadBaseAdr + (DiagVars.LogHeader.LogMemSize - DiagVars.LogMemToGet);// destination address
              StandardRequest.aData[4]        := DiagVars.BytesToGet$USINT;                   // length of data

              LastRequest := _ReadData;

#ifdef SAFETY_PROTOCOL_ANALYZER_ACTIVATED
  RecordFrame((#StandardRequest)$^DINT, 1);
#endif

              //copy SDO into write-buffer
              ToStdLib.MemCpy(dest := #p_Handle_SDO_Write^.SDOStructure, source := #StandardRequest, size := (sizeof(SDOHeader.StdHeader.CRC) + StandardRequest.SDOHeader.Len));

              //mark SDO data as valid
              p_Handle_SDO_Write^.us_Status := SAFETY_SDO_DATA_VALID;

              if ( pISafety^.udVersion >= 16#1001 ) then
                SAFETY_iPushSafetyTask();
              end_if;
            else
              UnsafeScheduler := UnsafeSchedulerNonPriorData;
            end_if;

//**********************************************************************************************************************************************************
          UnsafeSchedulerNonPriorData:

            // every 5 secs check for a new safety project inside the cpu
            if b_CheckCRC & ((ops.tAbsolute - ud_LastCrcCheck) > SBF_CRC_CHECK_TIME ) then

              SDORequestBuffer.StdHeader.CRC  := 0;                                                         // CRC is always 0 in Std communication
              SDORequestBuffer.StdHeader.Cmd  := SBF_SDO_COMMAND_READ;                                       // read command
              SDORequestBuffer.StdHeader.Typ  := SDO_STD;                                                   // standard frame type
              SDORequestBuffer.StdHeader.SeqNr:= StandardSeqNr OR 16#80;                                    // sequence number
              SDORequestBuffer.StdHeader.Len  := 4 + 4 + 1;                                                 // header + destination address + length of data
              SDORequestBuffer.ud_Address     := SBF_SDO_ADDRESS_CONFIG_DATA + SBF_SDO_OFFSET_CONFIG_CRC_ALL; // address of crc
              SDORequestBuffer.us_Length      := 4;                                                         // length of crc

              LastRequest := _GetCRC;

#ifdef SAFETY_PROTOCOL_ANALYZER_ACTIVATED
  RecordFrame((#SDORequestBuffer)$^DINT, 1);
#endif

              //copy SDO into write-buffer
              ToStdLib.MemCpy(dest := #p_Handle_SDO_Write^.SDOStructure, source := #SDORequestBuffer, size := (sizeof(SDOHeader.StdHeader.CRC) + SDORequestBuffer.StdHeader.Len));

              //mark SDO data as valid
              p_Handle_SDO_Write^.us_Status := SAFETY_SDO_DATA_VALID;

              if ( pISafety^.udVersion >= 16#1001 ) then
                SAFETY_iPushSafetyTask();
              end_if;

              ud_LastCrcCheck := ops.tAbsolute;

            // every 5 seconds write system time of plc to scp
            elsif b_SetSysTime & ((ops.tAbsolute - ud_LastSetSysTime) > SBF_SYSTIME_SET_TIME ) then

              if (LastRequest = _NoOpenRequest) & (p_Handle_SDO_Write^.us_Status = SAFETY_SDO_NO_DATA) then
                StandardRequest.SDOHeader.CRC  := 0;                               // CRC is always 0 in Std communication
                StandardRequest.SDOHeader.Cmd  := SBF_SDO_COMMAND_WRITE;           // read command
                StandardRequest.SDOHeader.Typ  := SDO_STD;                         // standard frame type
                StandardRequest.SDOHeader.SeqNr:= StandardSeqNr OR 16#80;          // sequence number
                StandardRequest.SDOHeader.Len  := 4 + 4 + 1 + sizeof(UDINT);       // header + destination address + length of data + size of data
                StandardRequest.aData[0]$UDINT := SBF_SDO_ADDRESS_FW_SYSTIME;      // address of system time safety firmware
                StandardRequest.aData[4]       := sizeof(UDINT);                   // length of data
                StandardRequest.aData[5]$UDINT := ToSigCLib.UnixTimeStampGet();    // system time of plc as unix timestamp

                LastRequest := _WriteSysTime;

                //copy SDO into write-buffer
                ToStdLib.MemCpy(dest := #p_Handle_SDO_Write^.SDOStructure, source := #StandardRequest, size := (sizeof(SDOHeader.StdHeader.CRC) + StandardRequest.SDOHeader.Len));

                //mark SDO data as valid
                p_Handle_SDO_Write^.us_Status := SAFETY_SDO_DATA_VALID;

                if ( pISafety^.udVersion >= 16#1001 ) then
                  SAFETY_iPushSafetyTask();
                end_if;

                ud_LastSetSysTime := ops.tAbsolute;
              end_if;

            else
              if RunState & us_SetBusReadyState = SetBusReadyFinished then
                // in operational (and SetbusReady is finished) also get unsafe-variables
                UnsafeScheduler := UnsafeSchedulerWriteData;
              else
                // not operational, we must skip the unsave vars
                UnsafeScheduler := UnsafeSchedulerDiagState;
                us_UnsafeSchedulerRun += 2;
              end_if;
            end_if;

//**********************************************************************************************************************************************************
          UnsafeSchedulerWriteData:

            if IsOptimizedCPU() then
              if ui_CntUnsafeInputs then
                // if we have finished checking through all variables the last time => check from beginning (otherwise the pointer is on the element where we have to continue)
                if pUnsafeInElement = NIL then
                  pUnsafeInElement := p_UnsafeInputsTable;
                end_if;

                // we check if we have to write any of the unsafe input variables (only until our message is full)
                UnsafeWrPackageNo := 0;
                BDINTWriteVars := 0; // limit number of bdint write variables to 3 to ensure constant load of firmware
                while pUnsafeInElement & (UnsafeWrPackageNo < SBF_MAX_UNSAFE_WRITE_PACKAGES) & (BDINTWriteVars < SBF_MAX_UNSAFE_BDINTS_PER_WRITE) do

                  // we have to check if we add this one
                  GotNewUnsafeValue := FALSE;

                  // if the type is normal we can read the actual value from the server
                  if pUnsafeInElement^.UnsafeType = NormalUnsafe then
                    // check if pointer to server is valid
                    if pUnsafeInElement^.ud_Thisp then
                      // get the actual value from the server
                      TmpVal := RD((pUnsafeInElement^.ud_Thisp)$^void);

                      // we remember to update this if it's necessary
                      GotNewUnsafeValue := TRUE;
                    else
                      if bd_LogOnceMarker.NoThisForUnsafeIn = FALSE then
                        bd_LogOnceMarker.NoThisForUnsafeIn := TRUE;
                        LogError("@0269 (SafetyBaseFSoE::CyWork) [SL] No thispointer available for Server of local unsafe input variable.");
                      end_if;
                    end_if;
                  elsif pUnsafeInElement^.UnsafeType = ExternalInput then
                    // check if we already have a valid value there
                    if pUnsafeInElement^.b_IsValid then
                      // get the actual value from the element
                      TmpVal := pUnsafeInElement^.sd_NewValue4External;

                      // we remember to update this if it's necessary
                      GotNewUnsafeValue := TRUE;
                    end_if;
                  else
                    if bd_LogOnceMarker.WrongUnsafeVarType = FALSE then
                      bd_LogOnceMarker.WrongUnsafeVarType := TRUE;
                      LogError("@026A (SafetyBaseFSoE::CyWork) [SL] Wrong unsafe variable type in unsafe input list.");
                    end_if;
                  end_if;

                  // if we have a new valid unsafe value => check if we have to send it
                  if GotNewUnsafeValue then
                    // if it hasn't been sent yet
                    if (pUnsafeInElement^.b_AlreadyTransmitted = FALSE) then
                      // remember that we sent this already
                      pUnsafeInElement^.b_AlreadyTransmitted := TRUE;

                      // add this one
                      AddUnsafePackage := TRUE;
                    elsif TmpVal <> pUnsafeInElement^.sd_OldValue then
                      // if there were any changes on this value

                      // add this one
                      AddUnsafePackage := TRUE;
                    else
                      // don't add this one
                      AddUnsafePackage := FALSE;
                    end_if;

                    // if it is ready to be added => add it to send buffer
                    if AddUnsafePackage then
                      // add a package to send
                      aUnsafeWrPackages[UnsafeWrPackageNo].ud_Address := pUnsafeInElement^.ud_Address;
                      aUnsafeWrPackages[UnsafeWrPackageNo].Value      := TmpVal;
                      UnsafeWrPackageNo += 1;

                      // if it has a bitmask it's an unsafe bdint input variable
                      if pUnsafeInElement^.BitMask then
                        BDINTWriteVars += 1;
                      end_if;

                      // remember the actual as old value
                      pUnsafeInElement^.sd_OldValue := TmpVal;
                    end_if;
                  end_if;

                  pUnsafeInElement := pUnsafeInElement^.pNext;
                end_while;

                if UnsafeWrPackageNo then
                  DataLen := UnsafeWrPackageNo * sizeof(UnsafeWritePackage);

                  StandardRequest.SDOHeader.Cmd                 := SBF_SDO_COMMAND_WRITE_VALUES;    // write values command
                  StandardRequest.SDOHeader.Typ                 := SDO_STD;                        // standard frame type
                  StandardRequest.SDOHeader.SeqNr               := StandardSeqNr OR 16#80;         // sequence number is in special area
                  StandardRequest.SDOHeader.Len                 := 4 + 4 + 1 + DataLen;            // header + destination address + length of data + data
                  StandardRequest.aData[0]                      := UnsafeWrPackageNo;              // number of packages
                  StandardRequest.aData[1]$UnsafeWritePackages  := aUnsafeWrPackages;              // packages

                  LastRequest := _WriteValues;

#ifdef SAFETY_PROTOCOL_ANALYZER_ACTIVATED
  RecordFrame((#StandardRequest)$^DINT, 1);
#endif

                  //copy SDO into write-buffer
                  ToStdLib.MemCpy(dest := #p_Handle_SDO_Write^.SDOStructure, source := #StandardRequest, size := (sizeof(SDOHeader.StdHeader.CRC) + StandardRequest.SDOHeader.Len));

                  //mark SDO data as valid
                  p_Handle_SDO_Write^.us_Status := SAFETY_SDO_DATA_VALID;

                  if ( pISafety^.udVersion >= 16#1001 ) then
                    SAFETY_iPushSafetyTask();
                  end_if;
                else
                  UnsafeScheduler := UnsafeSchedulerReadData;
                end_if;
              else
                UnsafeScheduler := UnsafeSchedulerReadData;
              end_if;
            else
              // on CSCP011 the SDO_COMMAND_WRITE_VALUES didn't exist
              if ui_CntUnsafeInputs & WriteFramesNeeded then
                // if writing is not active, check if it's necessary to activate it
                if (UnsafeWritingActive = FALSE) then
                  pUnsafeInElement := p_UnsafeInputsTable;

                  for i := 0 to (ui_CntUnsafeInputs - 1) do
                    if pUnsafeInElement^.ud_Thisp then
                      sd_retval := RD((pUnsafeInElement^.ud_Thisp)$^void);        // data
                      if pUnsafeInElement^.sd_OldValue <> sd_retval then
                        UnsafeWritingActive := TRUE;
                        pUnsafeInElement^.sd_OldValue := sd_retval;
                      end_if;
                    end_if;
                    pUnsafeInElement += sizeof(UnsafeIORoutingElement);
                  end_for;
                end_if;

                // check if writing is already active
                if UnsafeWritingActive then
                  // pointer to the right unsafe input
                  pUnsafeInElement := p_UnsafeInputsTable + (UnsafeWriteTransNr * MaxVarsPerWritePackage * sizeof(UnsafeIORoutingElement));

                  // get length of data we write
                  if (UnsafeWriteTransNr < (WriteFramesNeeded-1)) | ((ui_CntUnsafeInputs MOD MaxVarsPerWritePackage) = 0) then
                    DataLen := MaxVarsPerWritePackage * sizeof(DINT);
                  else
                    DataLen := (ui_CntUnsafeInputs MOD MaxVarsPerWritePackage)$USINT * sizeof(DINT);
                  end_if;

                  StandardRequest.SDOHeader.Cmd   := SBF_SDO_COMMAND_WRITE;                        // write command
                  StandardRequest.SDOHeader.Typ   := SDO_STD;                                     // standard frame type
                  StandardRequest.SDOHeader.SeqNr := StandardSeqNr OR 16#80;                      // sequence number is in special area
                  StandardRequest.SDOHeader.Len   := 4 + 4 + 1 + DataLen;                         // header + destination address + length of data + data
                  StandardRequest.aData[0]$UDINT  := pUnsafeInElement^.ud_Address;                // destination address
                  StandardRequest.aData[4]        := DataLen;                                     // length of data

                  // depending on length we do different number of server read-methods to get the data we write
                  for i := 0 to (DataLen/sizeof(DINT)) - 1 do
                    if pUnsafeInElement^.ud_Thisp then
                      StandardRequest.aData[5 + (i * sizeof(DINT))]$DINT := pUnsafeInElement^.sd_OldValue;
                    else
                      // this server doesn't exist in lasal => always send 0
                      StandardRequest.aData[5 + (i * sizeof(DINT))]$DINT := 0;
                    end_if;

                    pUnsafeInElement += sizeof(UnsafeIORoutingElement);
                  end_for;

                  LastRequest := _WriteValues;

#ifdef SAFETY_PROTOCOL_ANALYZER_ACTIVATED
  RecordFrame((#StandardRequest)$^DINT, 1);
#endif

                  //copy SDO into write-buffer
                  ToStdLib.MemCpy(dest := #p_Handle_SDO_Write^.SDOStructure, source := #StandardRequest, size := (sizeof(SDOHeader.StdHeader.CRC) + StandardRequest.SDOHeader.Len));

                  //mark SDO data as valid
                  p_Handle_SDO_Write^.us_Status := SAFETY_SDO_DATA_VALID;

                  if ( pISafety^.udVersion >= 16#1001 ) then
                    SAFETY_iPushSafetyTask();
                  end_if;
                else
                  UnsafeScheduler := UnsafeSchedulerReadData;
                end_if;
              else
                UnsafeScheduler := UnsafeSchedulerReadData;
              end_if;
            end_if;

//**********************************************************************************************************************************************************
          UnsafeSchedulerReadData:

            if ui_CntUnsafeOutputs & ReadFramesNeeded then
              //check, if buffer is empty and we got some unsafe data to get/set and crc check is finished
              if (UnsafeReadTransNr < ReadFramesNeeded) //then
               & ( ((UnsafeReadTransNr = 0) & ( ops.tAbsolute - LastUnsafeUpdate > ud_ServerUpdateTime ) ) | (UnsafeReadTransNr <> 0) )then
                // here we request directly the unsafe IOs

                // sequence number is in special area
                StandardRequest.SDOHeader.SeqNr := StandardSeqNr OR 16#80;

                // we get an output
                pUnsafeOutElement := p_UnsafeOutputsTable + (UnsafeReadTransNr * MaxVarsPerReadPackage * sizeof(UnsafeIORoutingElement));

                // get length of data we read
                if (UnsafeReadTransNr < (ReadFramesNeeded - 1)) | ((ui_CntUnsafeOutputs MOD MaxVarsPerReadPackage) = 0) then
                  UnsafeRdPackageNo := MaxVarsPerReadPackage;
                else
                  UnsafeRdPackageNo := (ui_CntUnsafeOutputs MOD MaxVarsPerReadPackage)$USINT;
                end_if;

                DataLen := UnsafeRdPackageNo * sizeof(DINT);

                // create buffer with addresses of values to read
                pHelpUnsafe := pUnsafeOutElement;
                for i := 0 to (UnsafeRdPackageNo-1) do
                  aUnsafeRdPackages[i] := pHelpUnsafe^.ud_Address;
                  pHelpUnsafe += sizeof(UnsafeIORoutingElement);
                end_for;

                StandardRequest.SDOHeader.Cmd               := SBF_SDO_COMMAND_READ_VALUES;                  // read values command
                StandardRequest.SDOHeader.Typ               := SDO_STD;                                     // standard frame type
                StandardRequest.SDOHeader.SeqNr             := StandardSeqNr OR 16#80;                      // sequence number is in special area
                StandardRequest.SDOHeader.Len               := 4 + 1 + DataLen;                             // header + size + length of data
                StandardRequest.aData[0]                    := UnsafeRdPackageNo;                           // number of values to get
                StandardRequest.aData[1]$UnsafeReadPackages := aUnsafeRdPackages;                           // read addresses

                LastRequest := _ReadValues;

#ifdef SAFETY_PROTOCOL_ANALYZER_ACTIVATED
  RecordFrame((#StandardRequest)$^DINT, 1);
#endif

                //copy SDO into write-buffer
                ToStdLib.MemCpy(dest := #p_Handle_SDO_Write^.SDOStructure, source := #StandardRequest, size := (sizeof(SDOHeader.StdHeader.CRC) + StandardRequest.SDOHeader.Len));

                //mark SDO data as valid
                p_Handle_SDO_Write^.us_Status := SAFETY_SDO_DATA_VALID;

                if ( pISafety^.udVersion >= 16#1001 ) then
                  SAFETY_iPushSafetyTask();
                end_if;

              elsif (UnsafeReadTransNr >= ReadFramesNeeded) then
                // We have finished all read data, go on with the next step
                UnsafeScheduler := UnsafeSchedulerDiagState;
                LastUnsafeUpdate := ops.tAbsolute;
                UnsafeReadTransNr := 0;
              else
                // time until read is not yet over - go on
                UnsafeScheduler := UnsafeSchedulerDiagState;
              end_if;
            else
              UnsafeScheduler := UnsafeSchedulerDiagState;
            end_if;

//**********************************************************************************************************************************************************
          UnsafeSchedulerDiagState:

            // get the diag state (on user demand)
            if DiagVars.UserWantsDiagState then

              // get state via SDO communication
              SDORequestBuffer.StdHeader.CRC  := 0;                                                   // CRC is always 0 in Std communication
              SDORequestBuffer.StdHeader.Cmd  := SBF_SDO_COMMAND_GET_STATE;                            // get-state command
              SDORequestBuffer.StdHeader.Typ  := SDO_STD;                                             // standard frame type
              SDORequestBuffer.StdHeader.SeqNr:= StandardSeqNr OR 16#80;                              // sequence number
              SDORequestBuffer.StdHeader.Len  := 4;                                                   // header
              SDORequestBuffer.ud_Address     := 0;
              SDORequestBuffer.us_Length      := 0;

              LastRequest := _DiagState;

#ifdef SAFETY_PROTOCOL_ANALYZER_ACTIVATED
  RecordFrame((#SDORequestBuffer)$^DINT, 1);
#endif

              //copy SDO into write-buffer
              ToStdLib.MemCpy(dest := #p_Handle_SDO_Write^.SDOStructure, source := #SDORequestBuffer, size := (sizeof(SDOHeader.StdHeader.CRC) + SDORequestBuffer.StdHeader.Len));

              //mark SDO data as valid
              p_Handle_SDO_Write^.us_Status := SAFETY_SDO_DATA_VALID;

              if ( pISafety^.udVersion >= 16#1001 ) then
                SAFETY_iPushSafetyTask();
              end_if;
            else
              UnsafeScheduler := UnsafeSchedulerDiagInfo;
            end_if;

//**********************************************************************************************************************************************************
            UnsafeSchedulerDiagInfo:

            // get the diag info (on user demand)
            if DiagVars.UserWantsDiagInfo then

              // get state via SDO communication
              StandardRequest.SDOHeader.CRC  := 0;                                                   // CRC is always 0 in Std communication
              StandardRequest.SDOHeader.Cmd  := SBF_SDO_COMMAND_GET_DIAG_INFO;                        // read command
              StandardRequest.SDOHeader.Typ  := SDO_STD;                                             // standard frame type
              StandardRequest.SDOHeader.SeqNr:= StandardSeqNr OR 16#80;                              // sequence number
              StandardRequest.SDOHeader.Len  := 4 + 1;                                               // header + µC-selection
              StandardRequest.aData[0] := DiagVars.ucChoiceDiagInfo;

              LastRequest := _DiagInfo;

#ifdef SAFETY_PROTOCOL_ANALYZER_ACTIVATED
  RecordFrame((#StandardRequest)$^DINT, 1);
#endif

              //copy SDO into write-buffer
              ToStdLib.MemCpy(dest := #p_Handle_SDO_Write^.SDOStructure, source := #StandardRequest, size := (sizeof(SDOHeader.StdHeader.CRC) + StandardRequest.SDOHeader.Len));

              //mark SDO data as valid
              p_Handle_SDO_Write^.us_Status := SAFETY_SDO_DATA_VALID;

              if ( pISafety^.udVersion >= 16#1001 ) then
                SAFETY_iPushSafetyTask();
              end_if;

            else

//              if SchedulerStepNo = 6 then
//                UnsafeScheduler := UnsafeSchedulerGetDiagVars;
//
//              elsif SchedulerStepNo = 7 then
//                UnsafeScheduler := UnsafeSchedulerGetRetryCounter;
//              end_if;
              UnsafeScheduler := UnsafeSchedulerGetRetryCounter;

            end_if;

//**********************************************************************************************************************************************************
          UnsafeSchedulerGetRetryCounter:

            //read out the retry counters every 10seconds
            if (b_RetryCounterAvailable) & (b_DisableSafetyRetryCnt = FALSE)
            & ((ops.tAbsolute - ud_RetryCntTimeMark) > SBF_RETRY_COUNTER_WAIT_TIME)  then

              SDORequestBuffer.StdHeader.CRC  := 0;                                                         // CRC is always 0 in Std communication
              SDORequestBuffer.StdHeader.Cmd  := SBF_SDO_COMMAND_READ;                                       // read command
              SDORequestBuffer.StdHeader.Typ  := SDO_STD;                                                   // standard frame type
              SDORequestBuffer.StdHeader.SeqNr:= StandardSeqNr OR 16#80;                                    // sequence number
              SDORequestBuffer.StdHeader.Len  := 4 + 4 + SBF_SDO_LENGTH_RETRY_COUNTER;                       // header + destination address + length of data
              SDORequestBuffer.ud_Address     := SBF_SDO_ADDRESS_RETRY_COUNTER;                              // address of retrycounter
              SDORequestBuffer.us_Length      := SBF_SDO_LENGTH_RETRY_COUNTER;                               // length of data

              LastRequest := _ReadRetryCounter;

#ifdef SAFETY_PROTOCOL_ANALYZER_ACTIVATED
  RecordFrame((#SDORequestBuffer)$^DINT, 1);
#endif

              //copy SDO into write-buffer
              ToStdLib.MemCpy(dest := #p_Handle_SDO_Write^.SDOStructure, source := #SDORequestBuffer, size := (sizeof(SDOHeader.StdHeader.CRC) + SDORequestBuffer.StdHeader.Len));

              //mark SDO data as valid
              p_Handle_SDO_Write^.us_Status := SAFETY_SDO_DATA_VALID;

              if ( pISafety^.udVersion >= 16#1001 ) then
                SAFETY_iPushSafetyTask();
              end_if;

              //reset timemark
              ud_RetryCntTimeMark := ops.tAbsolute;

            else
              UnsafeScheduler := UnsafeSchedulerChannelError;
            end_if;

//**********************************************************************************************************************************************************
          UnsafeSchedulerChannelError:

            if DiagVars.UserWantsErrorInfo  then
              SDORequestBuffer.StdHeader.CRC  := 0;                                                          // CRC is always 0 in Std communication
              SDORequestBuffer.StdHeader.Cmd  := SBF_SDO_COMMAND_READ;                                       // read command
              SDORequestBuffer.StdHeader.Typ  := SDO_STD;                                                    // standard frame type
              SDORequestBuffer.StdHeader.SeqNr:= StandardSeqNr OR 16#80;                                     // sequence number
              SDORequestBuffer.StdHeader.Len  := 4 + 4 + 1;                                                  // header + destination address + length of data
              SDORequestBuffer.ud_Address     := SBF_SDO_ADDRESS_ERROR_MEM;                                  // address of error memory
              SDORequestBuffer.us_Length      := SBF_SDO_LENGTH_ERROR_MESSAGE;                               // length of data (first byte contains number of following values + number of channels)

              if remainingPacketlength <> 0 then
                // set offset if more than one package
                SDORequestBuffer.ud_Address     := (SBF_SDO_ADDRESS_ERROR_MEM + actoffset);                  // address of error memory
                // set new length for next package
                if remainingPacketlength > SBF_SDO_LENGTH_ERROR_MESSAGE then
                  SDORequestBuffer.us_Length      := SBF_SDO_LENGTH_ERROR_MESSAGE;
                else
                  SDORequestBuffer.us_Length      := remainingPacketlength$USINT;
                end_if;
              end_if;

              LastRequest := _ErrorChannelInfo;

#ifdef SAFETY_PROTOCOL_ANALYZER_ACTIVATED
RecordFrame((#SDORequestBuffer)$^DINT, 1);
#endif

              //copy SDO into write-buffer
              ToStdLib.MemCpy(dest := #p_Handle_SDO_Write^.SDOStructure, source := #SDORequestBuffer, size := (sizeof(SDOHeader.StdHeader.CRC) + SDORequestBuffer.StdHeader.Len));

              //mark SDO data as valid
              p_Handle_SDO_Write^.us_Status := SAFETY_SDO_DATA_VALID;

              if ( pISafety^.udVersion >= 16#1001 ) then
                SAFETY_iPushSafetyTask();
              end_if;

              //reset timemark
              ud_RetryCntTimeMark := ops.tAbsolute;

            else
              UnsafeScheduler := UnsafeSchedulerGetFlexConNodeState;
            end_if;

//**********************************************************************************************************************************************************
          UnsafeSchedulerGetFlexConNodeState:

            // if there is a flexible constellation in the configuration and also an object placed and connected, we check the state regularly
            if (sFlexCon.FoundNodeInConfig) & ((ops.tAbsolute - sFlexCon.ud_LastNodeStateTimeStamp) > SBF_FLEX_CON_STATE_CHECK_TIME) then

              SDORequestBuffer.StdHeader.CRC  := 0;                                                         // CRC is always 0 in Std communication
              SDORequestBuffer.StdHeader.Cmd  := SBF_SDO_COMMAND_READ;                                      // read command
              SDORequestBuffer.StdHeader.Typ  := SDO_STD;                                                   // standard frame type
              SDORequestBuffer.StdHeader.SeqNr:= StandardSeqNr OR 16#80;                                    // sequence number
              SDORequestBuffer.StdHeader.Len  := 4 + 4 + sizeof(t_FlexConNodeState);                        // header + destination address + length of data
              SDORequestBuffer.ud_Address     := SBF_SDO_ADDRESS_FLEX_CON_NODE;                             // address of retrycounter
              SDORequestBuffer.us_Length      := sizeof(t_FlexConNodeState);                                // length of data

              LastRequest := _ReadFlexConNodeState;

#ifdef SAFETY_PROTOCOL_ANALYZER_ACTIVATED
  RecordFrame((#SDORequestBuffer)$^DINT, 1);
#endif

              //copy SDO into write-buffer
              ToStdLib.MemCpy(dest := #p_Handle_SDO_Write^.SDOStructure, source := #SDORequestBuffer, size := (sizeof(SDOHeader.StdHeader.CRC) + SDORequestBuffer.StdHeader.Len));

              //mark SDO data as valid
              p_Handle_SDO_Write^.us_Status := SAFETY_SDO_DATA_VALID;

              if ( pISafety^.udVersion >= 16#1001 ) then
                SAFETY_iPushSafetyTask();
              end_if;

              //reset timemark
              sFlexCon.ud_LastNodeStateTimeStamp := ops.tAbsolute;

            else
              UnsafeScheduler := UnsafeSchedulerGetFlexConHostState;
            end_if;

//**********************************************************************************************************************************************************
          UnsafeSchedulerGetFlexConHostState:

            // if there is a flexible constellation in the configuration and also an object placed and connected, we check the state regularly
            if (sFlexCon.FoundHostInConfig) & ((ops.tAbsolute - sFlexCon.ud_LastHostStateTimeStamp) > SBF_FLEX_CON_STATE_CHECK_TIME) then

              // calcuate max length
              us_SDO_length := SBF_SDO_MAX_LENGTH - (sizeof(SDOHeader) - sizeof(SDOHeader.SessId)) - sizeof(SDORespReadConfig.us_Returncode) - sizeof(SDORespReadConfig.us_Length);

              // if it's the first read of this run, read as much as possible (we don't know how many connections we have yet)
              if sFlexCon.LastHostState.CurrentReadOffset = 0 then
                // get maximum number of bytes
                DataLen := us_SDO_length;
              else
                // if we still need more or equal to max size
                if sFlexCon.LastHostState.BytesMissing >= us_SDO_length then
                  // get maximum number of bytes
                  DataLen := us_SDO_length;
                else
                  // otherwise it's the last package, so get the rest that is missing
                  DataLen := sFlexCon.LastHostState.BytesMissing$USINT;
                end_if;
              end_if;

              SDORequestBuffer.StdHeader.CRC  := 0;                                                                         // CRC is always 0 in Std communication
              SDORequestBuffer.StdHeader.Cmd  := SBF_SDO_COMMAND_READ;                                                      // read command
              SDORequestBuffer.StdHeader.Typ  := SDO_STD;                                                                   // standard frame type
              SDORequestBuffer.StdHeader.SeqNr:= StandardSeqNr OR 16#80;                                                    // sequence number
              SDORequestBuffer.StdHeader.Len  := 4 + 4 + sizeof(HDINT);                                                     // header + destination address + length of data
              SDORequestBuffer.ud_Address     := SBF_SDO_ADDRESS_FLEX_CON_HOST + sFlexCon.LastHostState.CurrentReadOffset;  // address of retrycounter
              SDORequestBuffer.us_Length      := DataLen;                                                                   // length of data

              // remember the length to check it when we receive the answer
              sFlexCon.LastHostState.LastRequestedLength := DataLen;

              LastRequest := _ReadFlexConHostState;

#ifdef SAFETY_PROTOCOL_ANALYZER_ACTIVATED
  RecordFrame((#SDORequestBuffer)$^DINT, 1);
#endif

              //copy SDO into write-buffer
              ToStdLib.MemCpy(dest := #p_Handle_SDO_Write^.SDOStructure, source := #SDORequestBuffer, size := (sizeof(SDOHeader.StdHeader.CRC) + SDORequestBuffer.StdHeader.Len));

              //mark SDO data as valid
              p_Handle_SDO_Write^.us_Status := SAFETY_SDO_DATA_VALID;

              if ( pISafety^.udVersion >= 16#1001 ) then
                SAFETY_iPushSafetyTask();
              end_if;

            else
              UnsafeScheduler := UnsafeSchedulerGetDiagVars;
            end_if;

//**********************************************************************************************************************************************************
        else
          if bd_LogOnceMarker.InvalidSchedulerState = FALSE then
            bd_LogOnceMarker.InvalidSchedulerState := TRUE;
            LogError("@026B (SafetyBaseFSoE::CyWork) [SL] Undefined Scheduler-State.");
          end_if;
        end_case;
      end_while;
    end_if;
  end_if;

  // at the first run we write all variables independent of any changes
  if RunState > OldRunState then
    SendAllUnsafeValues();
  end_if;
  OldRunState := RunState;

  state := READY;

//============================ Profiler start======================================================
#ifdef  DM_Profiler
  StopTimeMeasurement(usMode := DMTIME_CY);
#endif
//============================ Profiler end========================================================
END_FUNCTION

FUNCTION VIRTUAL SafetyBaseFSoE::GetConfiguration

END_FUNCTION

FUNCTION VIRTUAL SafetyBaseFSoE::SetSafetyState
  VAR_INPUT
    NewState 	: SafetyConfigStateType;
  END_VAR

  // use it locally => can also be forwarded in derivation
  SafetyState := NewState;

END_FUNCTION

FUNCTION VIRTUAL SafetyBaseFSoE::RefreshAsySrv
  // derive this
END_FUNCTION

FUNCTION VIRTUAL SafetyBaseFSoE::SetRetryCounter

  SafetyRetryCounter := -1;

END_FUNCTION

FUNCTION SafetyBaseFSoE::IsInCache
  VAR_INPUT
    ud_Address 	: UDINT;
    us_Length 	: USINT;
  END_VAR
  VAR_OUTPUT
    ItsInside 	: BOOL;
  END_VAR

  if CachedSize &
     (ud_Address >= CachedAddr) &
     ((ud_Address + us_Length) <= (CachedAddr + CachedSize)) then
    ItsInside := TRUE;
  else
    ItsInside := FALSE;
  end_if;

END_FUNCTION

FUNCTION SafetyBaseFSoE::AddToCache
  VAR_INPUT
    p_SDORequestBuffer 	: ^SDORequReadConfig;
    p_SDOResponseBuffer 	: ^SDORespReadConfig;
  END_VAR

  if p_SDORequestBuffer^.us_Length then
    CachedAddr := p_SDORequestBuffer^.ud_Address;
    CachedSize := p_SDORequestBuffer^.us_Length;
    _memcpy(ptr1:=#Cache, ptr2:=#p_SDOResponseBuffer^.ud_Data, cntr:=p_SDORequestBuffer^.us_Length);
  end_if;

END_FUNCTION

FUNCTION SafetyBaseFSoE::GetFSoEConnectionInfos
  VAR_INPUT
    p_SDORequestBuffer 	: ^SafetyBaseFSoE::SDORequReadConfig;
    p_SDOResponseBuffer 	: ^SafetyBaseFSoE::SDORespReadConfig;
  END_VAR
  VAR
    Address         : UDINT;
    Size            : USINT;
    sd_retval       : DINT;
    i               : UDINT;
    pActConnection  : ^t_FSoEConnectionDetails;
    TempRoutingInfo : t_FSoERoutingInfoElement;
    NextAddress     : UDINT;
  END_VAR
